// TIA Portal V19 export
// export: Created 2026-10-15T10:10:37.2525789Z, ExportSetting WithDefaults, DisplayName Totally Integrated Automation Portal, DisplayVersion V19, DisplayName TIA Portal Openness, DisplayVersion V19, DisplayName TIA Portal Version Control Interface, DisplayVersion V19, DisplayName STEP 7 Professional, DisplayVersion V19, DisplayName STEP 7 Safety, DisplayVersion V19, DisplayName WinCC Basic/Comfort/Advanced, DisplayVersion V19, DisplayName WinCC Unified, DisplayVersion V19
FUNCTION "ROLL_WriteOutputs" : Void   // FC37, SCL
{ S7_Optimized_Access := 'TRUE' }
VERSION : 0.1
// stored: AutoNumber true, IsIECCheckEnabled false, SetENOAutomatically false, UDAEnableTagReadback false
   VAR_TEMP
      enabled : Bool;
   END_VAR
BEGIN

   IF "ROLL_IO".PhysicalIoConfigured THEN
       #enabled := "ROLL_IO".PhysicalOutputsEnabled AND NOT "ROLL_IO".Simulation AND NOT "ROLL_IO".ConversionFault;
       "Tag__639276557961655014" := #enabled AND "ROLL_IO".Output[16, 0];
       "Tag__639276557961724830" := #enabled AND "ROLL_IO".Output[16, 1];
       "Tag__639276557961774695" := #enabled AND "ROLL_IO".Output[16, 2];
       "Tag__639276557961834550" := #enabled AND "ROLL_IO".Output[16, 3];
       "Tag__639276557961894385" := #enabled AND "ROLL_IO".Output[16, 4];
       "Tag__639276557961944242" := #enabled AND "ROLL_IO".Output[16, 5];
       "Tag__639276557962004083" := #enabled AND "ROLL_IO".Output[16, 6];
       "Tag__639276557962063929" := #enabled AND "ROLL_IO".Output[16, 7];
       "Tag__639276557962123762" := #enabled AND "ROLL_IO".Output[17, 0];
       "Tag__639276557962173628" := #enabled AND "ROLL_IO".Output[17, 1];
       "Tag__639276557962233470" := #enabled AND "ROLL_IO".Output[17, 2];
       "Tag__639276557962293353" := #enabled AND "ROLL_IO".Output[17, 3];
       "Tag__639276557962353158" := #enabled AND "ROLL_IO".Output[17, 4];
       "Tag__639276557962403014" := #enabled AND "ROLL_IO".Output[17, 5];
       "Tag__639276557962462907" := #enabled AND "ROLL_IO".Output[17, 6];
       "Tag__639276557962512720" := #enabled AND "ROLL_IO".Output[17, 7];
       "Tag__639276557962572561" := #enabled AND "ROLL_IO".Output[18, 0];
       "Tag__639276557962632401" := #enabled AND "ROLL_IO".Output[18, 1];
       "Tag__639276557962682267" := #enabled AND "ROLL_IO".Output[18, 2];
       "Tag__639276557962742107" := #enabled AND "ROLL_IO".Output[18, 3];
       "Tag__639276557962791974" := #enabled AND "ROLL_IO".Output[18, 4];
       "Tag__639276557962851816" := #enabled AND "ROLL_IO".Output[18, 5];
       "Tag__639276557962911653" := #enabled AND "ROLL_IO".Output[18, 6];
       "Tag__639276557962961520" := #enabled AND "ROLL_IO".Output[18, 7];
       "Tag__639276557963021363" := #enabled AND "ROLL_IO".Output[19, 0];
       "Tag__639276557963071237" := #enabled AND "ROLL_IO".Output[19, 1];
       "Tag__639276557963121101" := #enabled AND "ROLL_IO".Output[19, 2];
       "Tag__639276557963181309" := #enabled AND "ROLL_IO".Output[19, 3];
       "Tag__639276557963240774" := #enabled AND "ROLL_IO".Output[19, 4];
       "Tag__639276557963290937" := #enabled AND "ROLL_IO".Output[19, 5];
       "Tag__639276557963360463" := #enabled AND "ROLL_IO".Output[19, 6];
       "Tag__639276557963420293" := #enabled AND "ROLL_IO".Output[19, 7];
       "Tag__639276557963480133" := #enabled AND "ROLL_IO".Output[20, 0];
       "Tag__639276557963530002" := #enabled AND "ROLL_IO".Output[20, 1];
       "Tag__639276557963579865" := #enabled AND "ROLL_IO".Output[20, 2];
       "Tag__639276557963639838" := #enabled AND "ROLL_IO".Output[20, 3];
       "Tag__639276557963699546" := #enabled AND "ROLL_IO".Output[20, 4];
       "Tag__639276557963749412" := #enabled AND "ROLL_IO".Output[20, 5];
       "Tag__639276557963799286" := #enabled AND "ROLL_IO".Output[20, 6];
       "Tag__639276557963859119" := #enabled AND "ROLL_IO".Output[20, 7];
       "Tag__639276557963908985" := #enabled AND "ROLL_IO".Output[21, 0];
       "Tag__639276557963968826" := #enabled AND "ROLL_IO".Output[21, 1];
       "Tag__639276557964018692" := #enabled AND "ROLL_IO".Output[21, 2];
       "Tag__639276557964068878" := #enabled AND "ROLL_IO".Output[21, 3];
       "Tag__639276557964128400" := #enabled AND "ROLL_IO".Output[21, 4];
       "Tag__639276557964188239" := #enabled AND "ROLL_IO".Output[21, 5];
       "Tag__639276557964248077" := #enabled AND "ROLL_IO".Output[21, 6];
       "Tag__639276557964298411" := #enabled AND "ROLL_IO".Output[21, 7];
       "Tag__639276557964357785" := #enabled AND "ROLL_IO".Output[22, 0];
       "Tag__639276557964417947" := #enabled AND "ROLL_IO".Output[22, 1];
       "Tag__639276557964477465" := #enabled AND "ROLL_IO".Output[22, 2];
       "Tag__639276557964527497" := #enabled AND "ROLL_IO".Output[22, 3];
       "Tag__639276557964587312" := #enabled AND "ROLL_IO".Output[22, 4];
       "Tag__639276557964637070" := #enabled AND "ROLL_IO".Output[22, 5];
       "Tag__639276557964697149" := #enabled AND "ROLL_IO".Output[22, 6];
       "Tag__639276557964746745" := #enabled AND "ROLL_IO".Output[22, 7];
       "Tag__639276557964816574" := #enabled AND "ROLL_IO".Output[23, 0];
       "Tag__639276557964876412" := #enabled AND "ROLL_IO".Output[23, 1];
       "Tag__639276557964936239" := #enabled AND "ROLL_IO".Output[23, 2];
       "Tag__639276557964986111" := #enabled AND "ROLL_IO".Output[23, 3];
       "Tag__639276557965046275" := #enabled AND "ROLL_IO".Output[23, 4];
       "Tag__639276557965095821" := #enabled AND "ROLL_IO".Output[23, 5];
       "Tag__639276557965155664" := #enabled AND "ROLL_IO".Output[23, 6];
       "Tag__639276557965205527" := #enabled AND "ROLL_IO".Output[23, 7];
       "Tag__639276557965265365" := #enabled AND "ROLL_IO".Output[24, 0];
       "Tag__639276557965325265" := #enabled AND "ROLL_IO".Output[24, 1];
       "Tag__639276557965375063" := #enabled AND "ROLL_IO".Output[24, 2];
       "Tag__639276557965434904" := #enabled AND "ROLL_IO".Output[24, 3];
       "Tag__639276557965484769" := #enabled AND "ROLL_IO".Output[24, 4];
       "Tag__639276557965544610" := #enabled AND "ROLL_IO".Output[24, 5];
       "Tag__639276557965604458" := #enabled AND "ROLL_IO".Output[24, 6];
       "Tag__639276557965654714" := #enabled AND "ROLL_IO".Output[24, 7];
       "Tag__639276557965714166" := #enabled AND "ROLL_IO".Output[25, 0];
       "Tag__639276557965774008" := #enabled AND "ROLL_IO".Output[25, 1];
       "Tag__639276557965834033" := #enabled AND "ROLL_IO".Output[25, 2];
       "Tag__639276557965893680" := #enabled AND "ROLL_IO".Output[25, 3];
       "Tag__639276557965953516" := #enabled AND "ROLL_IO".Output[25, 4];
       "Tag__639276557966003383" := #enabled AND "ROLL_IO".Output[25, 5];
       "Tag__639276557966063222" := #enabled AND "ROLL_IO".Output[25, 6];
       "Tag__639276557966113089" := #enabled AND "ROLL_IO".Output[25, 7];
   END_IF;
END_FUNCTION
